Staubli VAL3: pickPlaceCylinder.pgx

program pickPlaceCylinder()
// Picks red cylinder from dispenser and places it in the assembling station.
begin
  putln("[2/4] Transferring red cylinder to station...")
  open(tLateral)

  // Safe joint transit to avoid wrist/elbow flip
  movej(jTransCylinder, tLateral, mNomSpeed)
  waitEndMove()

  // Pick from dispenser
  movej(pCylApproach, tLateral, mNomSpeed)
  waitEndMove()
  movel(pCylPick, tLateral, mInsertSpeed)
  waitEndMove()
  close(tLateral)

  movel(pCylApproach, tLateral, mNomSpeed)
  waitEndMove()

  // Place in assembling station
  movej(pAsmApproach, tLateral, mNomSpeed)
  waitEndMove()
  movel(pAsmCylinder, tLateral, mInsertSpeed)
  waitEndMove()
  open(tLateral)

  movel(pAsmApproach, tLateral, mNomSpeed)
  waitEndMove()
end
